(* IEC 61131-3 sources: plc_generation_empirical_study/datasets/packages/internal_v0_1/qualification_only/C04_E01_rising_edge_pulse, 1 file *)

(* ---- reference.st ---- *)
FUNCTION_BLOCK C04_E01_rising_edge_pulse
VAR_INPUT
    Signal : BOOL;
END_VAR
VAR_OUTPUT
    Pulse : BOOL;
END_VAR
VAR
    PrevSignal : BOOL := FALSE;
END_VAR

Pulse := Signal AND (NOT PrevSignal);
PrevSignal := Signal;

END_FUNCTION_BLOCK
